// TIA Portal V20 export
// export: Created 2026-10-20T12:44:01.7865471Z, ExportSetting WithDefaults, DisplayName Totally Integrated Automation Portal, DisplayVersion V20 Update 6, DisplayName TIA Portal Openness, DisplayVersion V20 Update 6, DisplayName TIA Portal Version Control Interface, DisplayVersion V20 Update 6, DisplayName SINAMICS Startdrive Advanced, DisplayVersion V20 SP1, DisplayName SINAMICS Startdrive G130, G150, S120, S150, SINAMICS MV, G220, S200, S210, DisplayVersion V20 SP1, DisplayName SINAMICS Startdrive G110M, G120, G120C, G120D, G120P, G115D, DisplayVersion V20 SP1, DisplayName STEP 7 Professional, DisplayVersion V20 Update 6, DisplayName STEP 7 Safety, DisplayVersion V20 Update 2, DisplayName WinCC Basic/Comfort/Advanced, DisplayVersion V20 Update 6, DisplayName WinCC Unified, DisplayVersion V20 Update 6
DATA_BLOCK "OPC_Control_FB_DB_5"   // DB333
VERSION : 0.1
// stored: AutoNumber true, DBAccessibleFromOPCUA true, InstanceOfName OPC_Control_FB, InstanceOfType FB
"OPC_Control_FB"
   // VAR_INPUT
   //    Id : UInt;
   //    All_In_Automatic : Bool;
   //    VTD_Error : Bool;
   //    OPC_Enable : Bool;
   //    Clear_OrderTable : Bool;
   // END_VAR
   // VAR_OUTPUT
   //    Error_ID : Word;
   // END_VAR
   // VAR
   //    Source_Location { ExternalAccessible := 'False'; ExternalVisible := 'False'; ExternalWritable := 'False'} : "ID_Decoded";
   //    Destination_Location { ExternalAccessible := 'False'; ExternalVisible := 'False'; ExternalWritable := 'False'} : "ID_Decoded";
   //    State_Main : UInt;
   //    State_VTD : UInt;
   //    State_Shuttle : UInt;
   //    State_CNV : UInt;
   //    T_Wait_Report_Done { S7_SetPoint := 'True'} : TON_TIME;
   // END_VAR
BEGIN
END_DATA_BLOCK
